(*
SPDX-FileCopyrightText: © 2026 Oleksandr Tiutyk <trofimich@gmail.com>
SPDX-License-Identifier: MIT
License: https://opensource.org/license/mit
*)

(*!
<summary>
Beckhoff EP1809_0021: 16-channel digital input EtherCAT Box (24 V DC, 3 ms filter, M8).
</summary>
<description>
Process image mapping structure for the EP1809_0021 EtherCAT Box IP67 module with 16 discrete inputs.
When used for I/O, link located fields or their containing buffers to the matching selected PDOs.
The record is not a packed wire buffer; compiler padding is not part of the device specification.
Unlinked/default values do not prove valid I/O. The caller evaluates bus/channel validity before use.
Use one owner task per instance and externally synchronize other access; multi-field snapshots are not atomic.
Copies store data without creating hardware links. Keep borrowed field references valid while consumers are bound.
This passive record performs no validation, synchronization, configuration or protocol advancement.
</description>
*)
TYPE EP1809_0021 :
STRUCT
	Ch01 AT %I* : BOOL;
	Ch02 AT %I* : BOOL;
	Ch03 AT %I* : BOOL;
	Ch04 AT %I* : BOOL;
	Ch05 AT %I* : BOOL;
	Ch06 AT %I* : BOOL;
	Ch07 AT %I* : BOOL;
	Ch08 AT %I* : BOOL;
	Ch09 AT %I* : BOOL;
	Ch10 AT %I* : BOOL;
	Ch11 AT %I* : BOOL;
	Ch12 AT %I* : BOOL;
	Ch13 AT %I* : BOOL;
	Ch14 AT %I* : BOOL;
	Ch15 AT %I* : BOOL;
	Ch16 AT %I* : BOOL;
END_STRUCT
END_TYPE

(* stored: Version 1.1.0.1, ProductVersion 3.1.4026.20
   DUT EP1809_0021: Id {bdb94bcc-3cdd-4a26-b0e6-56963e7d42dc} *)
